Staubli VAL3: simulate_UI.pgx

program simulate_UI()
  local bool l_bExit
begin

  do
    if util:sPage!="simulate"
      util:sPage="simulate"
      userPageBind("simulate","lbl2","innerHTML",sMsg,1,"r")
      userPageBindClick("simulate","img1",bCancel,true)
      userPage("simulate")
      delay(0.1)
    endIf
    sMsg=rs:sTrajStatus
    if bCancel
      bCancel=false
      l_bExit=true
    endIf


    delay(0)
  until l_bExit==true or taskStatus("simulate")==-1
  rs:bSimulate=false
  rs:bGOTO=false
  if taskStatus("simulate")>-1
    taskKill("simulate")
    resetMotion()
  endIf

end
